(* IEC 61131-3 sources: Lasal-MCP/examples/SampleSource/5_ClassInputOutputSolution/Stations/MachineControl/MachineControl/Class/AlarmBufferBase, 1 file *)

(* ---- AlarmBufferBase.st ---- *)
(*!
<Class
	Name               = "AlarmBufferBase"
	Revision           = "1.9"
	RealtimeTask       = "false"
	CyclicTask         = "false"
	DefCyclictime      = "50 ms"
	BackgroundTask     = "false"
	Sigmatek           = "true"
	OSInterface        = "false"
	HighPriority       = "false"
	Automatic          = "false"
	UpdateMode         = "Prescan"
	SharedCommandTable = "true"
	Objectsize         = "(536,120)"
	Comment            = "This class collects infomations about active alarms and provides this informations.&#13;&#10;It&apos;s possible to derive several methods to evaluate the extended alarm informations.&#13;&#10;&#13;&#10;IMPORTANT:&#13;&#10;The class is not compatible with the standard alarm classes.&#13;&#10;Must be used in combination with following classes:&#13;&#10;- AlarmOPMode0Para&#13;&#10;- AlarmOPMode1Para&#13;&#10;- AlarmOPMode2Para&#13;&#10;- AlarmOPMode3Para&#13;&#10;&#13;&#10;Not possible to use more than one object of this class in the project. The name of this object must be _AlarmXBuffer1.">
	<Channels>
		<Server Name="actOPMode" Visualized="true" Initialize="false" WriteProtected="true" Retentive="false" Comment="Server shows the actual operation mode."/>
		<Server Name="AlarmInfo" Visualized="true" Initialize="false" WriteProtected="true" Retentive="false" Comment="Server shows the actual AlarmInfo. In case one alarm with an active bit of the AlarmInfo is active, this bit is set within the server AlarmInfo.&#13;&#10;&#13;&#10;Call read-methode to show the value!"/>
		<Server Name="GroupAutomatic" Visualized="true" Initialize="false" WriteProtected="true" Retentive="false" Comment="Server shows the number of active alarms of the group OPMode_Automatic.&#13;&#10;&#13;&#10;Call read-methode to show the value!"/>
		<Server Name="GroupError" Visualized="true" Initialize="false" WriteProtected="true" Retentive="false" Comment="Server shows the number of active alarms of the group OPMode_Error.&#13;&#10;&#13;&#10;Call read-methode to show the value!"/>
		<Server Name="GroupHoming" Visualized="true" Initialize="false" WriteProtected="true" Retentive="false" Comment="Server shows the number of active alarms of the group OPMode_Homing.&#13;&#10;&#13;&#10;Call read-methode to show the value!"/>
		<Server Name="GroupInit" Visualized="true" Initialize="false" WriteProtected="true" Retentive="false" Comment="Server shows the number of active alarms of the group OPMode_Init.&#13;&#10;&#13;&#10;Call read-methode to show the value!"/>
		<Server Name="GroupManual" Visualized="true" Initialize="false" WriteProtected="true" Retentive="false" Comment="Server shows the number of active alarms of the group OPMode_Manual.&#13;&#10;&#13;&#10;Call read-methode to show the value!"/>
		<Server Name="GroupSemiAuto" Visualized="true" Initialize="false" WriteProtected="true" Retentive="false" Comment="Server shows the number of active alarms of the group OPMode_SemiAuto.&#13;&#10;&#13;&#10;Call read-methode to show the value!"/>
		<Server Name="GroupSetup" Visualized="true" Initialize="false" WriteProtected="true" Retentive="false" Comment="Server shows the number of active alarms of the group OPMode_Setup.&#13;&#10;&#13;&#10;Call read-methode to show the value!"/>
		<Server Name="GroupStop" Visualized="true" Initialize="false" WriteProtected="true" Retentive="false" Comment="Server shows the number of active alarms of the group OPMode_Stop.&#13;&#10;&#13;&#10;Call read-methode to show the value!"/>
		<Client Name="coOPModeConfig" Required="true" Internal="false"/>
		<Client Name="Parameter1" Required="false" Internal="false" Comment="The value of the connected server gets added to every alarm. In case nothing is connected, nothing is done.&#13;&#10;&#13;&#10;For example: &#13;&#10;- Alarm got 2 parameter =&gt; value of the connected server is stored in parameter 3.&#13;&#10;- Alarm got 3 parameter =&gt; value of the connected server is stored in parameter 4."/>
		<Client Name="Parameter2" Required="false" Internal="false" Comment="The value of the connected server gets added to every alarm. In case nothing is connected, nothing is done.&#13;&#10;&#13;&#10;For example: &#13;&#10;- Alarm got 2 parameter =&gt; value of the connected server is stored in parameter 3.&#13;&#10;- Alarm got 3 parameter =&gt; value of the connected server is stored in parameter 4."/>
	</Channels>
	<Dependencies>
		<Files>
			<File Path=".\Class\AlarmBufferBase\AlarmBufferBase.pdf"/>
			<File Path=".\Class\AlarmBufferBase\AlarmBufBase.h" Include="true"/>
		</Files>
	</Dependencies>
	<RevDoku>
		<Owner Company="Sigmatek"/>
		<Dokumentation Revision="1.9" Date="2019-12-18" Author="BurSte" Company="Sigmatek" Description="Bugfix:  since V1.8 the sum alarm bit field is not built correctly - corrected code (taken from V1.7)"/>
		<Dokumentation Revision="1.8" Date="2018-02-08" Author="SchMat" Company="Sigmatek" Description="use method ActionAlarmIntern for additional data handling to ensure multithreading"/>
		<Dokumentation Revision="1.7" Date="2017-05-09" Author="KaiAnd" Company="Sigmatek" Description="--&gt; Overwrite method Quit_AlarmAllEx() to count the alarm-quits&#13;&#10;--&gt; new global method GetAlarmQuitCnt() returns the counter of the alarm-quits for external use"/>
		<Dokumentation Revision="1.6" Date="2016-08-09" Author="ObeChr" Company="Sigmatek" Description="AlarmInfo from other stations can now be evaluated within this class."/>
		<Dokumentation Revision="1.4" Date="2016-03-23" Author="ObeChr" Company="Sigmatek" Description="Number of active alarms from other stations can now be evaluated within this class."/>
		<Dokumentation Revision="1.3" Date="2015-10-15" Author="HubChr" Company="Sigmatek" Description="Fixed issue with define MAX_ALARMPARA (no manual reconfiguration necessary anymore). Leaving the define at value 3 when using older versions could cause access exceptions."/>
		<Dokumentation Revision="1.2" Date="2015-07-09" Author="ObeChr" Company="Sigmatek" Description="Removed unnecessary Debugger Trace entry that was triggered on every error acknowledge."/>
		<Dokumentation Revision="1.1" Date="2015-06-10" Author="ObeChr" Company="Sigmatek" Description="+) Server actOPMode is now visualized.&#13;&#10;+) Methode AlarmQuit is now working."/>
		<Dokumentation Revision="1.0" Date="2015-06-01" Author="ObeChr" Company="Sigmatek" Description="First version of class to handle alarms in combination with OPModes."/>
	</RevDoku>
	<Network Name="AlarmBufferBase">
		<!-- List of Components in this network -->
		<Components>
			<Object
				Name       = "_base"
				Class      = "_AlarmXBuffer"
				Position   = "(218,120)"
				Visualized = "true">
				<Channels>
					<Server Name="ClassSvr"/>
					<Server Name="QuitAll"/>
					<Server Name="QuitAllEx"/>
					<Server Name="QuitGroup"/>
					<Server Name="QuitGroupEx"/>
					<Client Name="No" Value="64"/>
				</Channels>
			</Object>
		</Components>
		<Comments>
		</Comments>
		<!-- List of Connections in this network -->
		<Connections>
			<Connection Source="this.ClassSvr" Destination="_base.ClassSvr" Vertices="(690,210),(518,210),"/>
			<Connection Source="this.QuitAll" Destination="_base.QuitAll" Vertices="(690,270),(518,270),"/>
			<Connection Source="_base.No" Destination="this.No" Vertices="(218,210),(38,210),"/>
			<Connection Source="this.QuitGroup" Destination="_base.QuitGroup" Vertices="(690,330),(518,390),"/>
		</Connections>
		<!-- Headerfiles -->
		<Options>
		</Options>
	</Network>
</Class>
*)
#pragma using _AlarmXBuffer

AlarmBufferBase : CLASS
: _AlarmXBuffer
	TYPE
#pragma pack(push, 1)
	  t_s_OPMode : STRUCT  //! <Type Public="true" Name="t_s_OPMode"/>
	    udOPModeInit : UDINT;
	    udOPModeHoming : UDINT;
	    udOPModeStop : UDINT;
	    udOPModeSetup : UDINT;
	    udOPModeManual : UDINT;
	    udOPModeSemiAuto : UDINT;
	    udOPModeAutomatic : UDINT;
	    udOPModeError : UDINT;
	  END_STRUCT;
#pragma pack(pop)
#pragma pack(push, 1)
	  t_s_AlarmClient : STRUCT
	    pThis : ^AlarmStation;
	    sAlarmList : t_s_OPMode;
	    bdAlarmInfo : BDINT
	    [
	      1 Bit1,
	      2 Bit2,
	      3 Bit3,
	      4 Bit4,
	      5 Bit5,
	      6 Bit6,
	      7 Bit7,
	      8 Bit8,
	      9 Bit9,
	      10 Bit10,
	      11 Bit11,
	      12 Bit12,
	      13 Bit13,
	      14 Bit14,
	      15 Bit15,
	      16 Bit16,
	      17 Bit17,
	      18 Bit18,
	      19 Bit19,
	      20 Bit20,
	      21 Bit21,
	      22 Bit22,
	      23 Bit23,
	      24 Bit24,
	      25 Bit25,
	      26 Bit26,
	      27 Bit27,
	      28 Bit28,
	      29 Bit29,
	      30 Bit30,
	      31 Bit31,
	      32 Bit32,
	    ];
	  END_STRUCT;
#pragma pack(pop)
	END_TYPE
  //Servers:
	actOPMode 	: SvrChCmd_t_e_OPMode;
	GroupInit 	: SvrCh_UDINT;
	GroupHoming 	: SvrCh_UDINT;
	GroupStop 	: SvrCh_UDINT;
	GroupSetup 	: SvrCh_UDINT;
	GroupManual 	: SvrCh_UDINT;
	GroupSemiAuto 	: SvrCh_UDINT;
	GroupAutomatic 	: SvrCh_UDINT;
	GroupError 	: SvrCh_UDINT;
	AlarmInfo 	: SvrCh_BDINT;
  //Clients:
	coOPModeConfig 	: CltChCmd_OPModeConfigBase;
	Parameter1 	: CltCh_DINT;
	Parameter2 	: CltCh_DINT;
  //Variables:
		bdAlarmInfo : BDINT
		[
		  1 Bit1,
		  2 Bit2,
		  3 Bit3,
		  4 Bit4,
		  5 Bit5,
		  6 Bit6,
		  7 Bit7,
		  8 Bit8,
		  9 Bit9,
		  10 Bit10,
		  11 Bit11,
		  12 Bit12,
		  13 Bit13,
		  14 Bit14,
		  15 Bit15,
		  16 Bit16,
		  17 Bit17,
		  18 Bit18,
		  19 Bit19,
		  20 Bit20,
		  21 Bit21,
		  22 Bit22,
		  23 Bit23,
		  24 Bit24,
		  25 Bit25,
		  26 Bit26,
		  27 Bit27,
		  28 Bit28,
		  29 Bit29,
		  30 Bit30,
		  31 Bit31,
		  32 Bit32,
		];

		bdAlarmInfoStations : BDINT
		[
		  1 Bit1,
		  2 Bit2,
		  3 Bit3,
		  4 Bit4,
		  5 Bit5,
		  6 Bit6,
		  7 Bit7,
		  8 Bit8,
		  9 Bit9,
		  10 Bit10,
		  11 Bit11,
		  12 Bit12,
		  13 Bit13,
		  14 Bit14,
		  15 Bit15,
		  16 Bit16,
		  17 Bit17,
		  18 Bit18,
		  19 Bit19,
		  20 Bit20,
		  21 Bit21,
		  22 Bit22,
		  23 Bit23,
		  24 Bit24,
		  25 Bit25,
		  26 Bit26,
		  27 Bit27,
		  28 Bit28,
		  29 Bit29,
		  30 Bit30,
		  31 Bit31,
		  32 Bit32,
		];

		bsConfig : BSINT
		[
		  1 Parameter1Connected,
		  2 Parameter2Connected,
		  3 OPModeConfig,
		];

		eCommand 	: t_e_AlarmCmd;
		pOPMode 	: ^OPModeConfigBase::t_bd_OPMode;
		sAlarmInfo : ARRAY [0..31] OF UDINT;

		sAlarmStations : ARRAY [0..MAX_ALARMCLIENTS-1] OF t_s_AlarmClient;

		sOPModeAlarm 	: t_s_OPMode;
		sOPModeStations 	: t_s_OPMode;
		udAlarmClients 	: UDINT;
		cntQuit_AlarmAllEx 	: UDINT;
  //Functions:

	FUNCTION VIRTUAL GLOBAL Init;

	FUNCTION VIRTUAL Quit_AlarmAllEx
		VAR_OUTPUT
			retcode 	: BOOL;
		END_VAR;

	FUNCTION VIRTUAL GLOBAL RegisterAlarmXPara
		VAR_INPUT
			pThis 	: ^void;
			config 	: UDINT;
			group 	: UDINT;
			no 	: UDINT;
			paras 	: ^UDINT;
		END_VAR
		VAR_OUTPUT
			retcode 	: UDINT;
		END_VAR;

	FUNCTION VIRTUAL GLOBAL ActionAlarmIntern
		VAR_INPUT
			pThis 	: UDINT;
			config 	: UDINT;
			group 	: UDINT;
			state 	: DINT;
			parano 	: UDINT;
			ppara 	: ^DINT;
		END_VAR;

	FUNCTION VIRTUAL OPModeChange
		VAR_INPUT
			eActOPMode 	: t_e_OPMode;
			eNewOPMode 	: t_e_OPMode;
		END_VAR
		VAR_OUTPUT
			bOK 	: BOOL;
		END_VAR;

	FUNCTION VIRTUAL OPModeActive
		VAR_INPUT
			eActOPMode 	: t_e_OPMode;
		END_VAR
		VAR_OUTPUT
			eNewOPMode 	: t_e_OPMode;
		END_VAR;

	FUNCTION VIRTUAL AlarmActive
		VAR_INPUT
			udNo 	: UDINT;
			eOPMode 	: t_e_OPMode;
			bdInfo 	: BDINT;
		END_VAR;

	FUNCTION VIRTUAL AlarmInactive
		VAR_INPUT
			udNo 	: UDINT;
			eOPMode 	: t_e_OPMode;
			bdInfo 	: BDINT;
		END_VAR;

	FUNCTION VIRTUAL AlarmQuit
		VAR_INPUT
			udNo 	: UDINT;
		END_VAR;

	FUNCTION GLOBAL LoginAlarmClient
		VAR_INPUT
			pThis 	: ^AlarmStation;
		END_VAR
		VAR_OUTPUT
			bSuccessful 	: BOOL;
		END_VAR;
				//! <Function Comment="Within this methode the number of active alarms for each client gets determined." Name="AlarmStations"/>
	FUNCTION AlarmStations;

	FUNCTION GLOBAL GetAlarmQuitCnt
		VAR_OUTPUT
			RetVal 	: UDINT;
		END_VAR;

	FUNCTION VIRTUAL GLOBAL actOPMode::NewInst
		VAR_INPUT
			pPara 	: ^CmdStruct;
			pResult 	: ^results;
		END_VAR
		VAR_OUTPUT
			ret_code 	: iprStates;
		END_VAR;

	FUNCTION VIRTUAL GLOBAL GroupInit::Read
		VAR_OUTPUT
			output (EAX) 	: UDINT;
		END_VAR;

	FUNCTION VIRTUAL GLOBAL GroupHoming::Read
		VAR_OUTPUT
			output (EAX) 	: UDINT;
		END_VAR;

	FUNCTION VIRTUAL GLOBAL GroupStop::Read
		VAR_OUTPUT
			output (EAX) 	: UDINT;
		END_VAR;

	FUNCTION VIRTUAL GLOBAL GroupSetup::Read
		VAR_OUTPUT
			output (EAX) 	: UDINT;
		END_VAR;

	FUNCTION VIRTUAL GLOBAL GroupManual::Read
		VAR_OUTPUT
			output (EAX) 	: UDINT;
		END_VAR;

	FUNCTION VIRTUAL GLOBAL GroupSemiAuto::Read
		VAR_OUTPUT
			output (EAX) 	: UDINT;
		END_VAR;

	FUNCTION VIRTUAL GLOBAL GroupAutomatic::Read
		VAR_OUTPUT
			output (EAX) 	: UDINT;
		END_VAR;

	FUNCTION VIRTUAL GLOBAL GroupError::Read
		VAR_OUTPUT
			output (EAX) 	: UDINT;
		END_VAR;

	FUNCTION VIRTUAL GLOBAL AlarmInfo::Read
		VAR_OUTPUT
			output (EAX) 	: BDINT;
		END_VAR;
  //Tables:
	FUNCTION @STD
		VAR_OUTPUT
			ret_code	: CONFSTATES;
		END_VAR;
	FUNCTION GLOBAL TAB @CT_;
END_CLASS;

#pragma usingLtd OPModeConfigBase

#pragma usingLtd AlarmStation

FUNCTION VIRTUAL GLOBAL AlarmBufferBase::Init
VAR
	tmpSize : DINT;
END_VAR

  // Call base-class
  _AlarmXBuffer::Init();

  // last init-run
  if _FirstScan then

    // get maximum number of additional parameter
    tmpSize := MAX_ALARMPARA;

    // check size of additional parameter
    if tmpSize < 5 then
      TRACE_ERR("Define MAX_ALARMPARA in AlarmXBuffer.h must be at least 5 => otherwise memoryleak");
    end_if;

  end_if;

END_FUNCTION

FUNCTION VIRTUAL GLOBAL AlarmBufferBase::RegisterAlarmXPara
	VAR_INPUT
		pThis 	: ^void;
		config 	: UDINT;
		group 	: UDINT;
		no 	: UDINT;
		paras 	: ^UDINT;
	END_VAR
	VAR_OUTPUT
		retcode 	: UDINT;
	END_VAR
  VAR
  	tmpPara   : ^UDINT;
    tmpOPMode : t_e_OPMode;
  END_VAR

  // check if additional parameters are available
  if no >= 1 then

    // check OPMode
    //---------------------------------------------------------------------
    // check if configuration of pOPMode is already available
    if bsConfig.OPModeConfig = false then

      // check if client Parameter1 is connected
      if IsClientConnected(input := #Parameter1) then
        bsConfig.Parameter1Connected := true;
      end_if;

      // check if client Parameter2 is connected
      if IsClientConnected(input := #Parameter2) then
        bsConfig.Parameter2Connected := true;
      end_if;

      pOPMode := coOPModeConfig.GetModeConfig();

      // check if configuration is valid
      if pOPMode <> NIL then
        bsConfig.OPModeConfig := true;
      else
        TRACE_ERR("AlarmBufferBase::RegisterAlarmXPara(): no configuration of OPMode available");
      end_if;

    end_if;

    // check if configured OPMode is available
    if bsConfig.OPModeConfig = true then

      // get selected OPMode
      tmpOPMode := (paras + (no - 1) * sizeof(UDINT))^$t_e_OPMode;

      // check if OPMode is available
      case tmpOPMode of

        //---------------------------------------------

        OPMode_Init:
          if pOPMode^.bOPModeInit = false then
            TRACE_ERR("AlarmBufferBase::RegisterAlarmXPara() OPMode_Init: invalid OPMode-configuration of alarm detected");
          end_if;

        //---------------------------------------------

        OPMode_Homing:
          if pOPMode^.bOPModeHoming = false then
            TRACE_ERR("AlarmBufferBase::RegisterAlarmXPara() OPMode_Homing: invalid OPMode-configuration of alarm detected");
          end_if;

        OPMode_Stop:
          if pOPMode^.bOPModeStop = false then
            TRACE_ERR("AlarmBufferBase::RegisterAlarmXPara() OPMode_Stop: invalid OPMode-configuration of alarm detected");
          end_if;

        //---------------------------------------------

        OPMode_Setup:
          if pOPMode^.bOPModeSetup = false then
            TRACE_ERR("AlarmBufferBase::RegisterAlarmXPara() OPMode_Setup: invalid OPMode-configuration of alarm detected");
          end_if;

        //---------------------------------------------

        OPMode_Manual:
          if pOPMode^.bOPModeManual = false then
            TRACE_ERR("AlarmBufferBase::RegisterAlarmXPara() OPMode_Manual: invalid OPMode-configuration of alarm detected");
          end_if;

        //---------------------------------------------

        OPMode_SemiAuto:
          if pOPMode^.bOPModeSemiAuto = false then
            TRACE_ERR("AlarmBufferBase::RegisterAlarmXPara() OPMode_SemiAuto: invalid OPMode-configuration of alarm detected");
          end_if;

        //---------------------------------------------

        OPMode_Automatic:
          if pOPMode^.bOPModeAutomatic = false then
            TRACE_ERR("AlarmBufferBase::RegisterAlarmXPara() OPMode_Automatic: invalid OPMode-configuration of alarm detected");
          end_if;

        //---------------------------------------------

        OPMode_Error:
          if pOPMode^.bOPModeError = false then
            TRACE_ERR("AlarmBufferBase::RegisterAlarmXPara() OPMode_Error: invalid OPMode-configuration of alarm detected");
          end_if;

        //---------------------------------------------

        else
          TRACE_ERR("AlarmBufferBase::RegisterAlarmXPara(): invalid operationmode detected");
      end_case;

    end_if;

    no -= 1;

    // Add Lasal ID of Parameter1 + Parameter2
    //---------------------------------------------------------------------
    // necessary, because the lse-kernel determines the configuration of
    // this connected dataserver (unit,...) Used to get the correct
    // formatting if the value is displayed on the screen.

    tmpPara := paras + no * sizeof(DINT);

    // check if Parameter 1 is connected
    if bsConfig.Parameter1Connected then
      tmpPara^ := (Parameter1.pCH)$UDINT;
      tmpPara += sizeof(DINT);
      no += 1;
    end_if;

    // check if Parameter 2 is connected
    if bsConfig.Parameter2Connected then
      tmpPara^ := (Parameter2.pCH)$UDINT;
      no += 1;
    end_if;

  else
    TRACE_ERR("AlarmBufferBase::RegisterAlarmXPara(): unkown alarm object detected");
  end_if;

  // call base class to login alarm
  //---------------------------------------------------------------------
  retcode := _AlarmXBuffer::RegisterAlarmXPara( pThis   := pThis,
                                                config  := config,
                                                group   := group,
                                                no      := no,
                                                paras   := paras);

END_FUNCTION

FUNCTION VIRTUAL GLOBAL AlarmBufferBase::actOPMode::NewInst
	VAR_INPUT
		pPara 	: ^CmdStruct;
		pResult 	: ^Results;
	END_VAR
	VAR_OUTPUT
		ret_code 	: IprStates;
	END_VAR

  // check input parameter
  if pPara = NIL | pResult = NIL then
    ret_code := ERROR;
    return;
  end_if;

  //*****************************************************************************
  //** CHECK TYPE OF COMMAND                                                   **
  //*****************************************************************************

  case pPara^.uiCmd$t_e_AlarmCmd of

    // Methode for active OPMode
    //***************************************************************************
    Cmd_OPModeActive:

      // set length of result
      pResult^.uiLng := sizeof(t_e_OPMode);

      // call methode for active OPMode
      pResult^.aData[0]$t_e_OPMode := OPModeActive(eActOPMode := pPara^.aPara[0]$t_e_OPMode);

      ret_code := READY;

    // Methode for changing OPMode
    //***************************************************************************
    Cmd_OPModeChange:

      // set length of result
      pResult^.uiLng := sizeof(BOOL);

      // call methode for changing OPMode
      pResult^.aData[0] := OPModeChange(eActOPMode  := pPara^.aPara[0]$t_e_OPMode,
                                        eNewOPMode  := pPara^.aPara[1]$t_e_OPMode);

      ret_code := READY;

    // new OPMode aktive
    //**************************************************************************
    Cmd_ActOPMode:

      actOPMode := pPara^.aPara[0]$t_e_OPMode;
      ret_code := READY;

     // unknown command
     //***************************************************************************
     else
      TRACE_ERR("AlarmBufferBase::actOPMode::NewInst(): unknown command");
      ret_code := ERROR;

  end_case;

END_FUNCTION

FUNCTION VIRTUAL AlarmBufferBase::OPModeChange
	VAR_INPUT
		eActOPMode 	: t_e_OPMode;
		eNewOPMode 	: t_e_OPMode;
	END_VAR
	VAR_OUTPUT
		bOK 	: BOOL;
	END_VAR

  // init returncode
  bOK := true;

  // get alarms from other stations
  AlarmStations();

  //*****************************************************************************
  //** DEPENDING ON THE NEW OPMODE DIFFERENT ALARMS GET CHECKED                **
  //*****************************************************************************

  case eNewOPMode of

    //***************************************************************************

    OPMode_Init:
      // nothing happens because of an alarm

    //***************************************************************************

    OPMode_Homing:

      // if at least one alarm is active => change to OPMode_Error
      if sOPModeAlarm.udOPModeHoming |
         sOPModeStations.udOPModeHoming then
        bOK := false;
      end_if;

    //***************************************************************************

    OPMode_Manual:

      // if at least one alarm is active => change to OPMode_Error
      if sOPModeAlarm.udOPModeManual |
         sOPModeStations.udOPModeManual then
        bOK := false;
      end_if;

    //***************************************************************************

    OPMode_SemiAuto:

      // if at least one alarm is active => change to OPMode_Error
      if sOPModeAlarm.udOPModeManual | sOPModeAlarm.udOPModeSemiAuto |
         sOPModeStations.udOPModeManual | sOPModeStations.udOPModeSemiAuto then
        bOK := false;
      end_if;

    //***************************************************************************

    OPMode_Automatic:

      // if at least one alarm is active => change to OPMode_Error
      if sOPModeAlarm.udOPModeManual | sOPModeAlarm.udOPModeSemiAuto | sOPModeAlarm.udOPModeAutomatic |
         sOPModeStations.udOPModeManual | sOPModeStations.udOPModeSemiAuto | sOPModeStations.udOPModeAutomatic  then
        bOK := false;
      end_if;

    //***************************************************************************

    OPMode_Error:

    //***************************************************************************

    else
      TRACE_ERR("AlarmBufferBase::OPModeChange(): not supported OPMode");

  end_case;

END_FUNCTION

FUNCTION VIRTUAL AlarmBufferBase::OPModeActive
	VAR_INPUT
		eActOPMode 	: t_e_OPMode;
	END_VAR
	VAR_OUTPUT
		eNewOPMode 	: t_e_OPMode;
	END_VAR

  // init returncode
  eNewOPMode := eActOPMode;

  // get alarms from other stations
  AlarmStations();

  //*****************************************************************************
  //** DEPENDING ON THE OPMODE DIFFERENT ALARMS GET CHECKED                    **
  //*****************************************************************************

  case eActOPMode of

    //***************************************************************************

    OPMode_Init:
      // nothing happens because of an alarm

    //***************************************************************************

    OPMode_Homing:

      // if at least one alarm is active => change to OPMode_Error
      if sOPModeAlarm.udOPModeHoming |
         sOPModeStations.udOPModeHoming then
        eNewOPMode := OPMode_Error;
      end_if;

    //***************************************************************************

    OPMode_Manual:

      // if at least one alarm is active => change to OPMode_Error
      if sOPModeAlarm.udOPModeManual |
         sOPModeStations.udOPModeManual then
        eNewOPMode := OPMode_Error;
      end_if;

    //***************************************************************************

    OPMode_SemiAuto:

      // if at least one alarm for OPMode_Manual is active => change to OPMode_Error
      if sOPModeAlarm.udOPModeManual |
         sOPModeStations.udOPModeManual then
        eNewOPMode := OPMode_Error;

      // if at least one alarm for OPMode_SemiAuto is active => change to OPMode_Manual
      elsif sOPModeAlarm.udOPModeSemiAuto |
            sOPModeStations.udOPModeSemiAuto then
        eNewOPMode := OPMode_Manual;
      end_if;

    //***************************************************************************

    OPMode_Automatic:

      // if at least one alarm for OPMode_Manual is active => change to OPMode_Error
      if sOPModeAlarm.udOPModeManual |
         sOPModeStations.udOPModeManual then
        eNewOPMode := OPMode_Error;
      // if at least one alarm for OPMode_SemiAuto is active => change to OPMode_Manual
      elsif sOPModeAlarm.udOPModeSemiAuto |
            sOPModeStations.udOPModeSemiAuto then
        eNewOPMode := OPMode_Manual;
      // if at least one alarm for OPMode_Automatic is active => change to OPMode_SemiAuto
      elsif sOPModeAlarm.udOPModeAutomatic |
            sOPModeStations.udOPModeAutomatic then
        eNewOPMode := OPMode_SemiAuto;
      end_if;

    //***************************************************************************

    OPMode_Error:

    //***************************************************************************

    else
      TRACE_ERR("AlarmBufferBase::OPModeActive(): not supported OPMode");

  end_case;

END_FUNCTION

FUNCTION GLOBAL AlarmBufferBase::LoginAlarmClient
	VAR_INPUT
		pThis 	: ^AlarmStation;
	END_VAR
	VAR_OUTPUT
		bSuccessful 	: BOOL;
	END_VAR

  // check input-parameter
  if pThis = NIL then
    bSuccessful := false;
    return;

  // check limits of array
  elsif udAlarmClients >= sizeof(sAlarmStations) / sizeof(sAlarmStations[0]) then
    bSuccessful := false;
    return;

  end_if;

  // save pointer
  sAlarmStations[udAlarmClients].pThis := pThis;
  udAlarmClients += 1;

  // set returncode
  bSuccessful := true;

END_FUNCTION

FUNCTION AlarmBufferBase::AlarmStations
  VAR
    tmpCounter  : UDINT;
    tmpObject   : ^AlarmStation;
  END_VAR

  // check if stations are available
  if udAlarmClients then

    bdAlarmInfoStations := 0;
    _memset(#sOPModeStations, 0, sizeof(sOPModeStations));

    // loop to get alarminformation from all connected client
    for tmpCounter := 0 to udAlarmClients - 1 do

      // get pointer to object
      tmpObject := sAlarmStations[tmpCounter].pThis;

      // check if pointer is valid
      if tmpObject <> NIL then

        // call methode to fetch information
        if tmpObject^.GetAlarms(pAlarms     := #sAlarmStations[tmpCounter].sAlarmList,
                                pAlarmInfo  := (#sAlarmStations[tmpCounter].bdAlarmInfo)$^BDINT) = true then

          // calculate sum of all clients
          sOPModeStations.udOPModeInit       += sAlarmStations[tmpCounter].sAlarmList.udOPModeInit;
          sOPModeStations.udOPModeHoming     += sAlarmStations[tmpCounter].sAlarmList.udOPModeHoming;
          sOPModeStations.udOPModeStop       += sAlarmStations[tmpCounter].sAlarmList.udOPModeStop;
          sOPModeStations.udOPModeSetup      += sAlarmStations[tmpCounter].sAlarmList.udOPModeSetup;
          sOPModeStations.udOPModeManual     += sAlarmStations[tmpCounter].sAlarmList.udOPModeManual;
          sOPModeStations.udOPModeSemiAuto   += sAlarmStations[tmpCounter].sAlarmList.udOPModeSemiAuto;
          sOPModeStations.udOPModeAutomatic  += sAlarmStations[tmpCounter].sAlarmList.udOPModeAutomatic;
          sOPModeStations.udOPModeError      += sAlarmStations[tmpCounter].sAlarmList.udOPModeError;

          // alarminfo from all clients
          bdAlarmInfoStations := bdAlarmInfoStations OR sAlarmStations[tmpCounter].bdAlarmInfo;

        else
          TRACE_ERR("AlarmBufferBase::CheckClient(): failed to fetch alarminformation from client");
        end_if;

      end_if;

    end_for;

  end_if;

END_FUNCTION

#pragma warning (disable: 73);
FUNCTION VIRTUAL AlarmBufferBase::AlarmActive
	VAR_INPUT
		udNo 	: UDINT;
		eOPMode 	: t_e_OPMode;
		bdInfo 	: BDINT;
	END_VAR
#pragma warning (default: 73);

END_FUNCTION

#pragma warning (disable: 73);
FUNCTION VIRTUAL AlarmBufferBase::AlarmInactive
	VAR_INPUT
		udNo 	: UDINT;
		eOPMode 	: t_e_OPMode;
		bdInfo 	: BDINT;
	END_VAR
#pragma warning (default: 73);

END_FUNCTION

#pragma warning (disable: 73);
FUNCTION VIRTUAL AlarmBufferBase::AlarmQuit
	VAR_INPUT
		udNo 	: UDINT;
	END_VAR
#pragma warning (default: 73);

END_FUNCTION

FUNCTION VIRTUAL GLOBAL AlarmBufferBase::GroupInit::Read
	VAR_OUTPUT
		output (EAX) 	: UDINT;
	END_VAR

  GroupInit := sOPModeAlarm.udOPModeInit;
	output := GroupInit;

END_FUNCTION

FUNCTION VIRTUAL GLOBAL AlarmBufferBase::GroupHoming::Read
	VAR_OUTPUT
		output (EAX) 	: UDINT;
	END_VAR

  GroupHoming := sOPModeAlarm.udOPModeHoming;
	output := GroupHoming;

END_FUNCTION

FUNCTION VIRTUAL GLOBAL AlarmBufferBase::GroupStop::Read
	VAR_OUTPUT
		output (EAX) 	: UDINT;
	END_VAR

  GroupStop := sOPModeAlarm.udOPModeStop;
	output := GroupStop;

END_FUNCTION

FUNCTION VIRTUAL GLOBAL AlarmBufferBase::GroupSetup::Read
	VAR_OUTPUT
		output (EAX) 	: UDINT;
	END_VAR

  GroupSetup := sOPModeAlarm.udOPModeSetup;
	output := GroupSetup;

END_FUNCTION

FUNCTION VIRTUAL GLOBAL AlarmBufferBase::GroupManual::Read
	VAR_OUTPUT
		output (EAX) 	: UDINT;
	END_VAR

  GroupManual := sOPModeAlarm.udOPModeManual;
	output := GroupManual;

END_FUNCTION

FUNCTION VIRTUAL GLOBAL AlarmBufferBase::GroupSemiAuto::Read
	VAR_OUTPUT
		output (EAX) 	: UDINT;
	END_VAR

  GroupSemiAuto := sOPModeAlarm.udOPModeSemiAuto;
	output := GroupSemiAuto;

END_FUNCTION

FUNCTION VIRTUAL GLOBAL AlarmBufferBase::GroupAutomatic::Read
	VAR_OUTPUT
		output (EAX) 	: UDINT;
	END_VAR

  GroupAutomatic := sOPModeAlarm.udOPModeAutomatic;
	output := GroupAutomatic;

END_FUNCTION

FUNCTION VIRTUAL GLOBAL AlarmBufferBase::GroupError::Read
	VAR_OUTPUT
		output (EAX) 	: UDINT;
	END_VAR

  GroupError := sOPModeAlarm.udOPModeError;
	output := GroupError;

END_FUNCTION

FUNCTION VIRTUAL GLOBAL AlarmBufferBase::AlarmInfo::Read
	VAR_OUTPUT
		output (EAX) 	: BDINT;
	END_VAR

  AlarmInfo := bdAlarmInfo;
	output := AlarmInfo;

END_FUNCTION

FUNCTION GLOBAL AlarmBufferBase::GetAlarmQuitCnt
	VAR_OUTPUT
		RetVal 	: UDINT;
	END_VAR

  RetVal := cntQuit_AlarmAllEx;

END_FUNCTION

FUNCTION VIRTUAL AlarmBufferBase::Quit_AlarmAllEx
	VAR_OUTPUT
		retcode 	: BOOL;
	END_VAR

  retCode := _AlarmXBuffer::Quit_AlarmAllEx();

  cntQuit_AlarmAllEx += 1;

END_FUNCTION

FUNCTION VIRTUAL GLOBAL AlarmBufferBase::ActionAlarmIntern
	VAR_INPUT
		pThis 	: UDINT;
		config 	: UDINT;
		group 	: UDINT;
		state 	: DINT;
		parano 	: UDINT;
		ppara 	: ^DINT;
	END_VAR
  VAR
  	tmpPara       : ^DINT;
    tmpValue      : SINT;
    tmpInfo       : BDINT;
    tmpMask       : BDINT;
    tmpAlarmInfo  : BDINT;
    tmpCounter    : USINT;
    tmpOPMode     : t_e_OPMode;
  END_VAR

  // check if additional parameters are available
  if parano >= 2 then

    // get parameters of alarm
    tmpOPMode := ((ppara + (parano - 2) * sizeof(DINT))^)$t_e_OPMode;
    tmpInfo   := ((ppara + (parano - 1) * sizeof(DINT))^)$BDINT;

    // count alarm for each OPMode
    //---------------------------------------------------------------------
    // alarm active
    if state > 0 then // HubChr v1.4 changed from "state = TRUE"
      tmpValue := 1;
    // alarm inacitve
    elsif state = false then
      tmpValue := -1;
    else
      tmpValue := 0;
    end_if;

    case tmpOPMode of

      OPMode_Init:
        sOPModeAlarm.udOPModeInit$DINT       += tmpValue;

      OPMode_Homing:
        sOPModeAlarm.udOPModeHoming$DINT     += tmpValue;

      OPMode_Stop:
        sOPModeAlarm.udOPModeStop$DINT       += tmpValue;

      OPMode_Setup:
        sOPModeAlarm.udOPModeSetup$DINT      += tmpValue;

      OPMode_Manual:
        sOPModeAlarm.udOPModeManual$DINT     += tmpValue;

      OPMode_SemiAuto:
        sOPModeAlarm.udOPModeSemiAuto$DINT   += tmpValue;

      OPMode_Automatic:
        sOPModeAlarm.udOPModeAutomatic$DINT  += tmpValue;

      OPMode_Error:
        sOPModeAlarm.udOPModeError$DINT      += tmpValue;

    else
      TRACE_ERR("AlarmBufferBase::ActionAlarm(): unkown operationmode detected");
    end_case;

    // check alarminfo
    //---------------------------------------------------------------------

    // reset alarminfo
    tmpAlarmInfo := 0;

    // evaluate each bit
    for tmpCounter := 0 to 31 do

      // build mask
      tmpMask := 2#1 SHL tmpCounter;

//v1.9 BruSte: Error Correction - with this Code some old AlarmInfos could be lost!
//      // check if bit is set
//      if tmpInfo AND tmpMask then
//
//        sAlarmInfo[tmpCounter]$DINT += tmpValue;
//
//        if sAlarmInfo[tmpCounter] then
//          tmpAlarmInfo := tmpAlarmInfo OR tmpMask;
//        end_if;
//
//      end_if;

//v1.9 BurSte: properly working old code from version v1.7

      // check if bit is set
      if tmpInfo AND tmpMask then
        sAlarmInfo[tmpCounter]$DINT += tmpValue;
      end_if;

      if sAlarmInfo[tmpCounter] then
        tmpAlarmInfo := tmpAlarmInfo OR tmpMask;
      end_if;

    end_for;

    // sum of all bits
    bdAlarmInfo := tmpAlarmInfo;

    // call user-methods
    //---------------------------------------------------------------------
    // alarm active
    if state > 0 then // HubChr v1.4 changed from "state = TRUE"
      AlarmActive(udNo    := config,
                  eOPMode := tmpOPMode,
                  bdInfo  := tmpInfo);
    // alarm inacitve
    elsif state = false then
      AlarmInactive(udNo    := config,
                    eOPMode := tmpOPMode,
                    bdInfo  := tmpInfo);
    elsif state <> -1 then
      TRACE_ERR("AlarmBufferBase::ActionAlarm(): unknown alarm state detected");
    end_if;

    // add Parameter 1 + Parameter 2
    //---------------------------------------------------------------------
    // get pointer behind the alarmparameter
    // the two parameter at the beginning are OPMode + AlarmInfo
    tmpPara := ppara + (parano - 2) * sizeof(DINT);

    // add parameter to alarm
    if bsConfig.Parameter1Connected then
      Parameter1  := Parameter1.Read();
      tmpPara^    := Parameter1;
      tmpPara     += sizeof(DINT);
    else
      parano -= 1;
    end_if;

    // add parameter to alarm
    if bsConfig.Parameter2Connected then
      Parameter2  := Parameter2.Read();
      tmpPara^    := Parameter2;
    else
      parano -= 1;
    end_if;

  elsif state <> -1 then
    TRACE_ERR("AlarmBufferBase::ActionAlarm(): unkown alarm object detected");
  end_if;

  // alarm quit
  if state = -1 then
    AlarmQuit(udNo    := config);
  end_if;

  // save alarm in AlarmBufferBase
  //---------------------------------------------------------------------
  _AlarmXBuffer::ActionAlarmIntern(pThis, config, group, state, parano, ppara);

END_FUNCTION
